FUNCTION F_DeadZone : REAL
(*
Function used to calculate dead zone.

Constructor: 		Patryk Panylo
Company:		E. Riexinger GmbH
Date:			03.06.2014
Version:			1.00

Date:			Revision:		Who:				Comment
dd.mm.yyyy		x.xx			Initials			comment

*)

VAR_INPUT
	(* Enummerations *)

	(* Variables *)
	lrInSignal								:LREAL;							(* Input signal *)
	lrDeadZone							:LREAL;							(* Dead zone *)

	(* References *)

	(* Interfaces *)

	(* Instances *)

END_VAR
VAR
	(* Enummerations *)

	(* Variables *)

	(* References *)

	(* Interfaces *)

	(* Instances *)

END_VAR


IF ABS(lrInSignal) > lrDeadZone
THEN
	F_DeadZone := lrInSignal;
ELSE
	F_DeadZone := 0.0;
END_IF;

END_FUNCTION

(* stored: Version 1.1.0.1, ProductVersion 3.1.4024.15
   POU F_DeadZone: Id {1148b447-6c19-41ca-b4fd-f4ad7fcd8dc5}, SpecialFunc None *)
